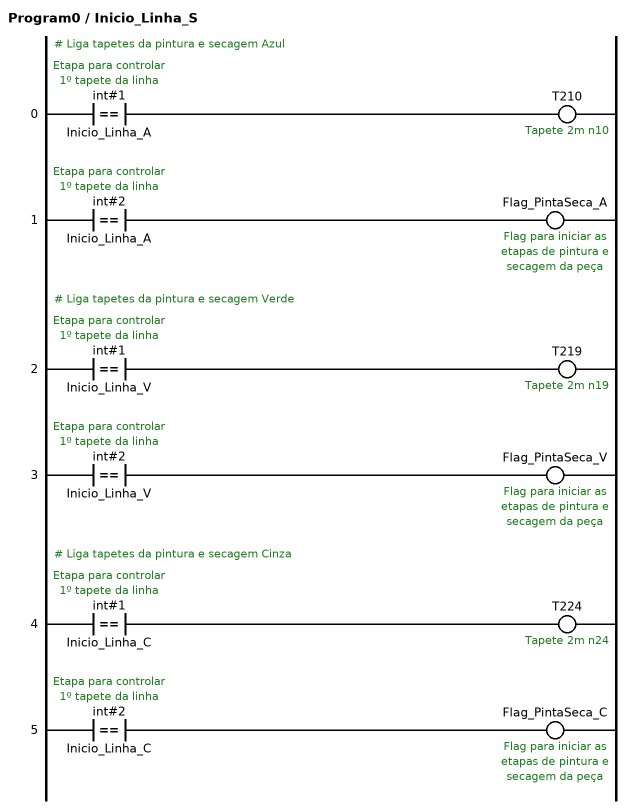
(* [picture p96: Program0 / Inicio_Linha_S, rungs 0-5] *)
(* Rung 0: # Liga tapetes da pintura e secagem Azul *)
T210 := int#1 = Inicio_Linha_A;
(* Rung 1 *)
Flag_PintaSeca_A := int#2 = Inicio_Linha_A;
(* Rung 2: # Liga tapetes da pintura e secagem Verde *)
T219 := int#1 = Inicio_Linha_V;
(* Rung 3 *)
Flag_PintaSeca_V := int#2 = Inicio_Linha_V;
(* Rung 4: # Liga tapetes da pintura e secagem Cinza *)
T224 := int#1 = Inicio_Linha_C;
(* Rung 5 *)
Flag_PintaSeca_C := int#2 = Inicio_Linha_C;

(* Section Pinta_Seca_E: ladder, written here as Structured Text *)

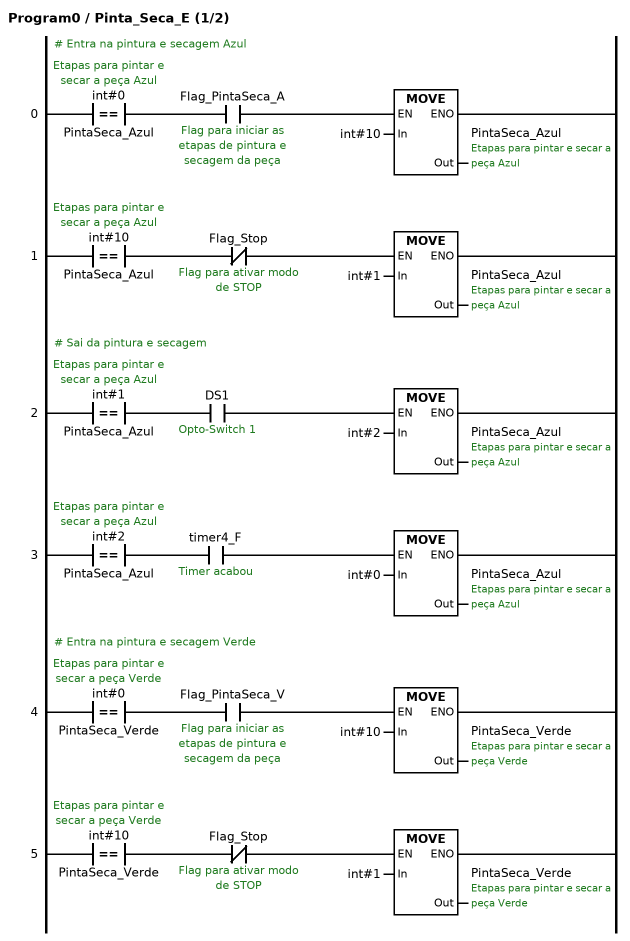
(* Rung 0: # Entra na pintura e secagem Azul *)
IF (int#0 = PintaSeca_Azul) AND Flag_PintaSeca_A THEN PintaSeca_Azul := int#10; END_IF;
(* Rung 1 *)
IF (int#10 = PintaSeca_Azul) AND NOT Flag_Stop THEN PintaSeca_Azul := int#1; END_IF;
(* Rung 2: # Sai da pintura e secagem *)
IF (int#1 = PintaSeca_Azul) AND DS1 THEN PintaSeca_Azul := int#2; END_IF;
(* Rung 3 *)
IF (int#2 = PintaSeca_Azul) AND timer4_F THEN PintaSeca_Azul := int#0; END_IF;
(* Rung 4: # Entra na pintura e secagem Verde *)
IF (int#0 = PintaSeca_Verde) AND Flag_PintaSeca_V THEN PintaSeca_Verde := int#10; END_IF;
(* Rung 5 *)
IF (int#10 = PintaSeca_Verde) AND NOT Flag_Stop THEN PintaSeca_Verde := int#1; END_IF;

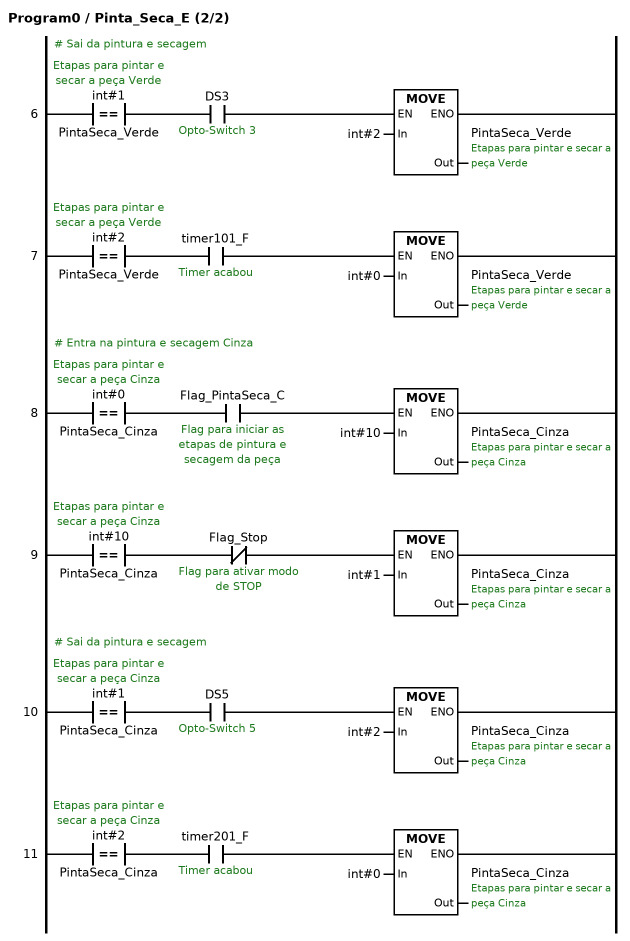
(* Rung 6: # Sai da pintura e secagem *)
IF (int#1 = PintaSeca_Verde) AND DS3 THEN PintaSeca_Verde := int#2; END_IF;
(* Rung 7 *)
IF (int#2 = PintaSeca_Verde) AND timer101_F THEN PintaSeca_Verde := int#0; END_IF;
(* Rung 8: # Entra na pintura e secagem Cinza *)
IF (int#0 = PintaSeca_Cinza) AND Flag_PintaSeca_C THEN PintaSeca_Cinza := int#10; END_IF;
(* Rung 9 *)
IF (int#10 = PintaSeca_Cinza) AND NOT Flag_Stop THEN PintaSeca_Cinza := int#1; END_IF;
(* Rung 10: # Sai da pintura e secagem *)
IF (int#1 = PintaSeca_Cinza) AND DS5 THEN PintaSeca_Cinza := int#2; END_IF;
(* Rung 11 *)
IF (int#2 = PintaSeca_Cinza) AND timer201_F THEN PintaSeca_Cinza := int#0; END_IF;

(* Section Pinta_Seca_S: ladder, written here as Structured Text *)

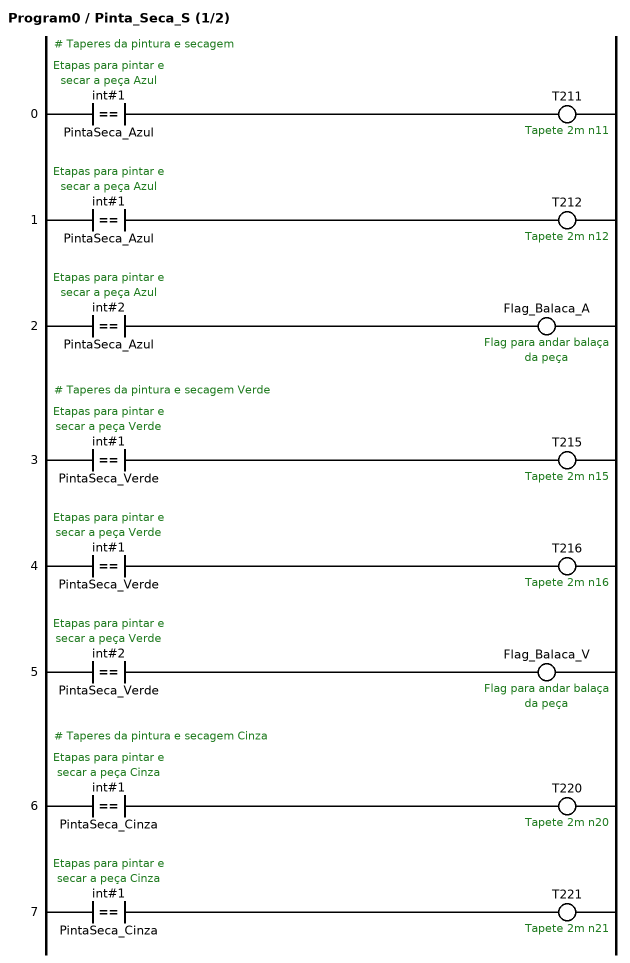
(* Rung 0: # Taperes da pintura e secagem *)
T211 := int#1 = PintaSeca_Azul;
(* Rung 1 *)
T212 := int#1 = PintaSeca_Azul;
(* Rung 2 *)
Flag_Balaca_A := int#2 = PintaSeca_Azul;
(* Rung 3: # Taperes da pintura e secagem Verde *)
T215 := int#1 = PintaSeca_Verde;
(* Rung 4 *)
T216 := int#1 = PintaSeca_Verde;
(* Rung 5 *)
Flag_Balaca_V := int#2 = PintaSeca_Verde;
(* Rung 6: # Taperes da pintura e secagem Cinza *)
T220 := int#1 = PintaSeca_Cinza;
(* Rung 7 *)
T221 := int#1 = PintaSeca_Cinza;

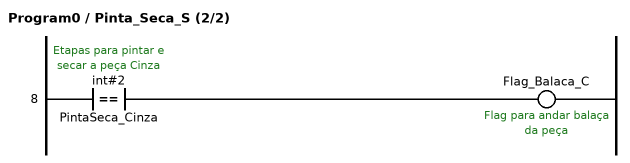
(* Rung 8 *)
Flag_Balaca_C := int#2 = PintaSeca_Cinza;

(* Section Balaca_E: ladder, written here as Structured Text *)

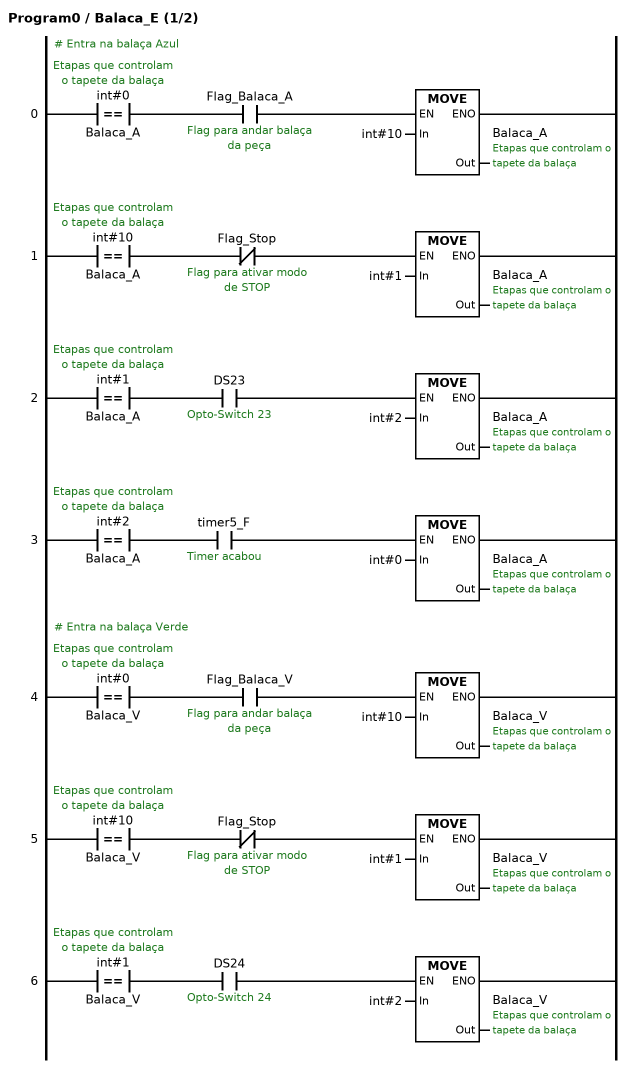
(* Rung 0: # Entra na balaça Azul *)
IF (int#0 = Balaca_A) AND Flag_Balaca_A THEN Balaca_A := int#10; END_IF;
(* Rung 1 *)
IF (int#10 = Balaca_A) AND NOT Flag_Stop THEN Balaca_A := int#1; END_IF;
(* Rung 2 *)
IF (int#1 = Balaca_A) AND DS23 THEN Balaca_A := int#2; END_IF;
(* Rung 3 *)
IF (int#2 = Balaca_A) AND timer5_F THEN Balaca_A := int#0; END_IF;
(* Rung 4: # Entra na balaça Verde *)
IF (int#0 = Balaca_V) AND Flag_Balaca_V THEN Balaca_V := int#10; END_IF;
(* Rung 5 *)
IF (int#10 = Balaca_V) AND NOT Flag_Stop THEN Balaca_V := int#1; END_IF;
(* Rung 6 *)
IF (int#1 = Balaca_V) AND DS24 THEN Balaca_V := int#2; END_IF;

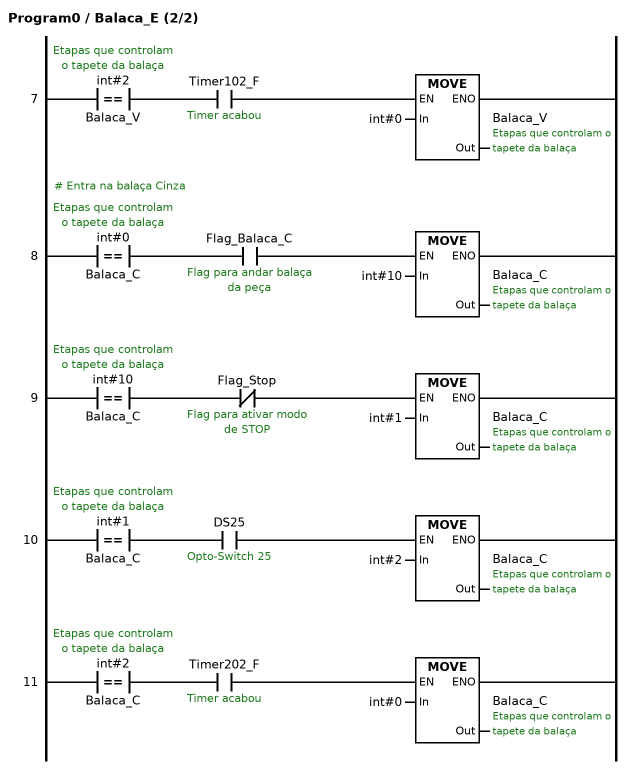
(* Rung 7 *)
IF (int#2 = Balaca_V) AND Timer102_F THEN Balaca_V := int#0; END_IF;
(* Rung 8: # Entra na balaça Cinza *)
IF (int#0 = Balaca_C) AND Flag_Balaca_C THEN Balaca_C := int#10; END_IF;
(* Rung 9 *)
IF (int#10 = Balaca_C) AND NOT Flag_Stop THEN Balaca_C := int#1; END_IF;
(* Rung 10 *)
IF (int#1 = Balaca_C) AND DS25 THEN Balaca_C := int#2; END_IF;
(* Rung 11 *)
IF (int#2 = Balaca_C) AND Timer202_F THEN Balaca_C := int#0; END_IF;

(* Section Balaca_S: ladder, written here as Structured Text *)

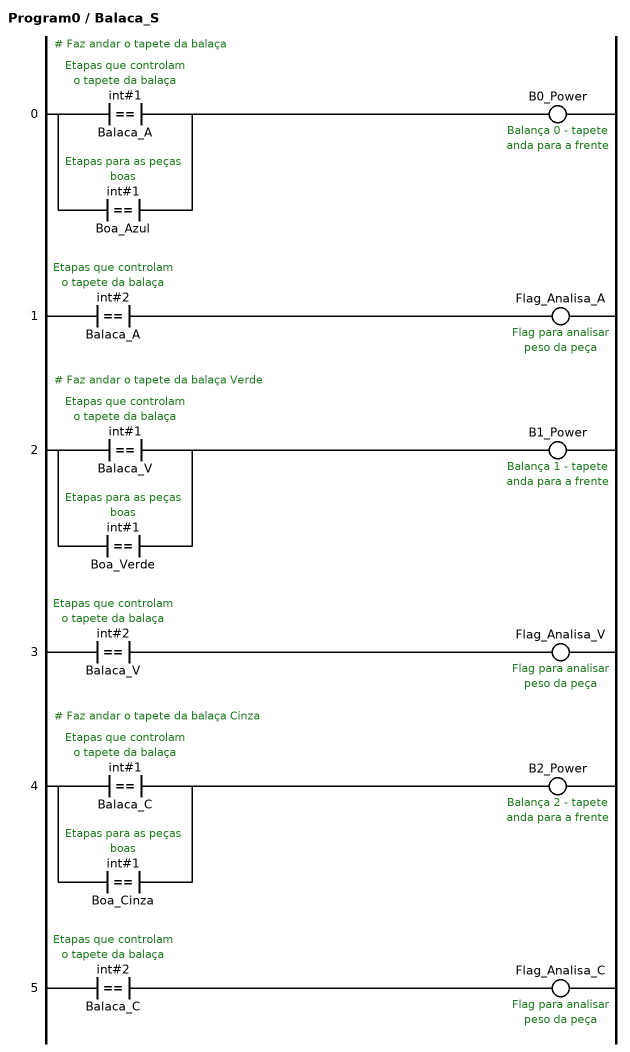
(* Rung 0: # Faz andar o tapete da balaça *)
B0_Power := (int#1 = Balaca_A) OR (int#1 = Boa_Azul);
(* Rung 1 *)
Flag_Analisa_A := int#2 = Balaca_A;
(* Rung 2: # Faz andar o tapete da balaça Verde *)
B1_Power := (int#1 = Balaca_V) OR (int#1 = Boa_Verde);
(* Rung 3 *)
Flag_Analisa_V := int#2 = Balaca_V;
(* Rung 4: # Faz andar o tapete da balaça Cinza *)
B2_Power := (int#1 = Balaca_C) OR (int#1 = Boa_Cinza);
(* Rung 5 *)
Flag_Analisa_C := int#2 = Balaca_C;

(* Section Analisa_Pesos_E: ladder, written here as Structured Text *)

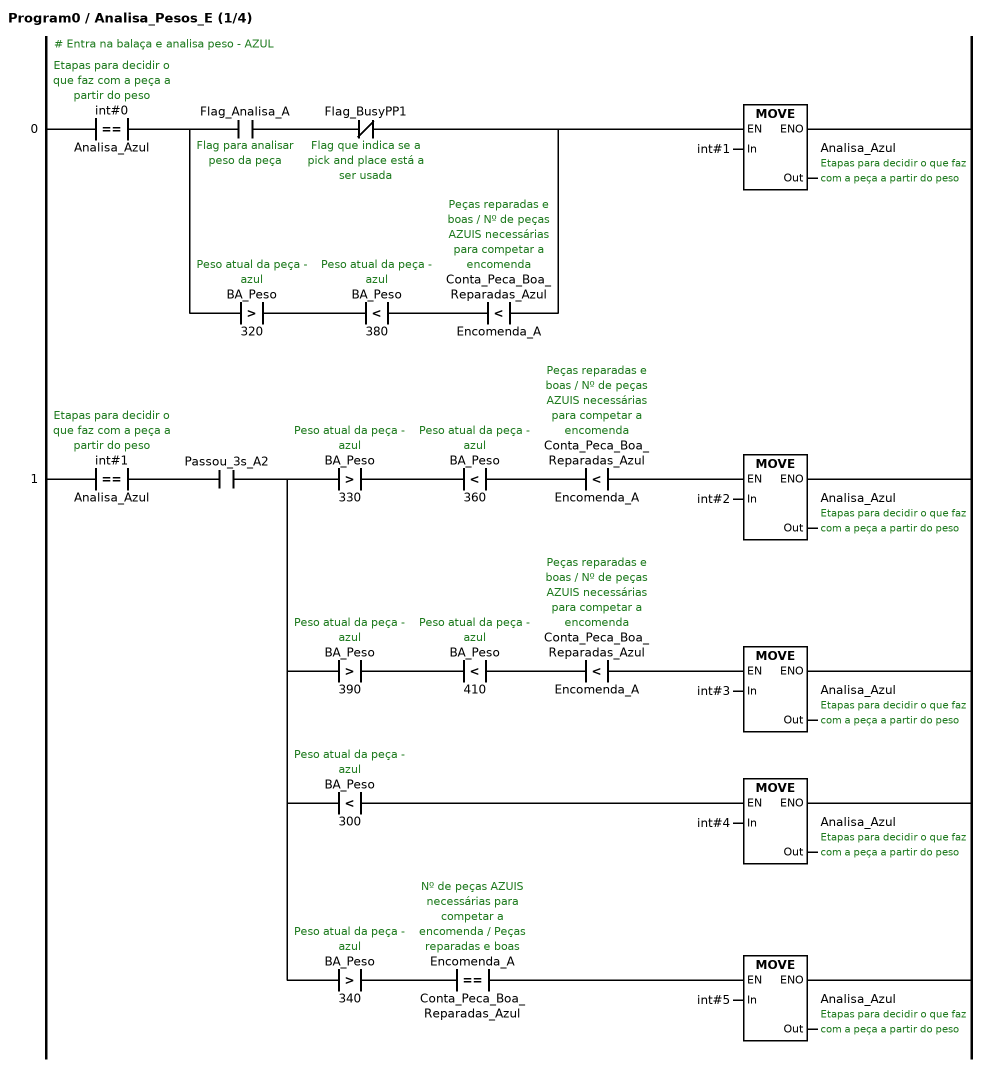
(* Rung 0: # Entra na balaça e analisa peso - AZUL *)
IF (int#0 = Analisa_Azul) AND ((Flag_Analisa_A AND NOT Flag_BusyPP1) OR ((BA_Peso > 320) AND (BA_Peso < 380) AND (Conta_Peca_Boa_Reparadas_Azul < Encomenda_A))) THEN
    Analisa_Azul := int#1;
END_IF;
(* Rung 1 *)
_p32 := (int#1 = Analisa_Azul) AND Passou_3s_A2;
IF (int#1 = Analisa_Azul) AND Passou_3s_A2 AND (BA_Peso > 330) AND (BA_Peso < 360) AND (Conta_Peca_Boa_Reparadas_Azul < Encomenda_A) THEN
    Analisa_Azul := int#2;
END_IF;
IF _p32 AND (BA_Peso > 390) AND (BA_Peso < 410) AND (Conta_Peca_Boa_Reparadas_Azul < Encomenda_A) THEN
    Analisa_Azul := int#3;
END_IF;
IF _p32 AND (BA_Peso < 300) THEN Analisa_Azul := int#4; END_IF;
IF _p32 AND (BA_Peso > 340) AND (Encomenda_A = Conta_Peca_Boa_Reparadas_Azul) THEN
    Analisa_Azul := int#5;
END_IF;

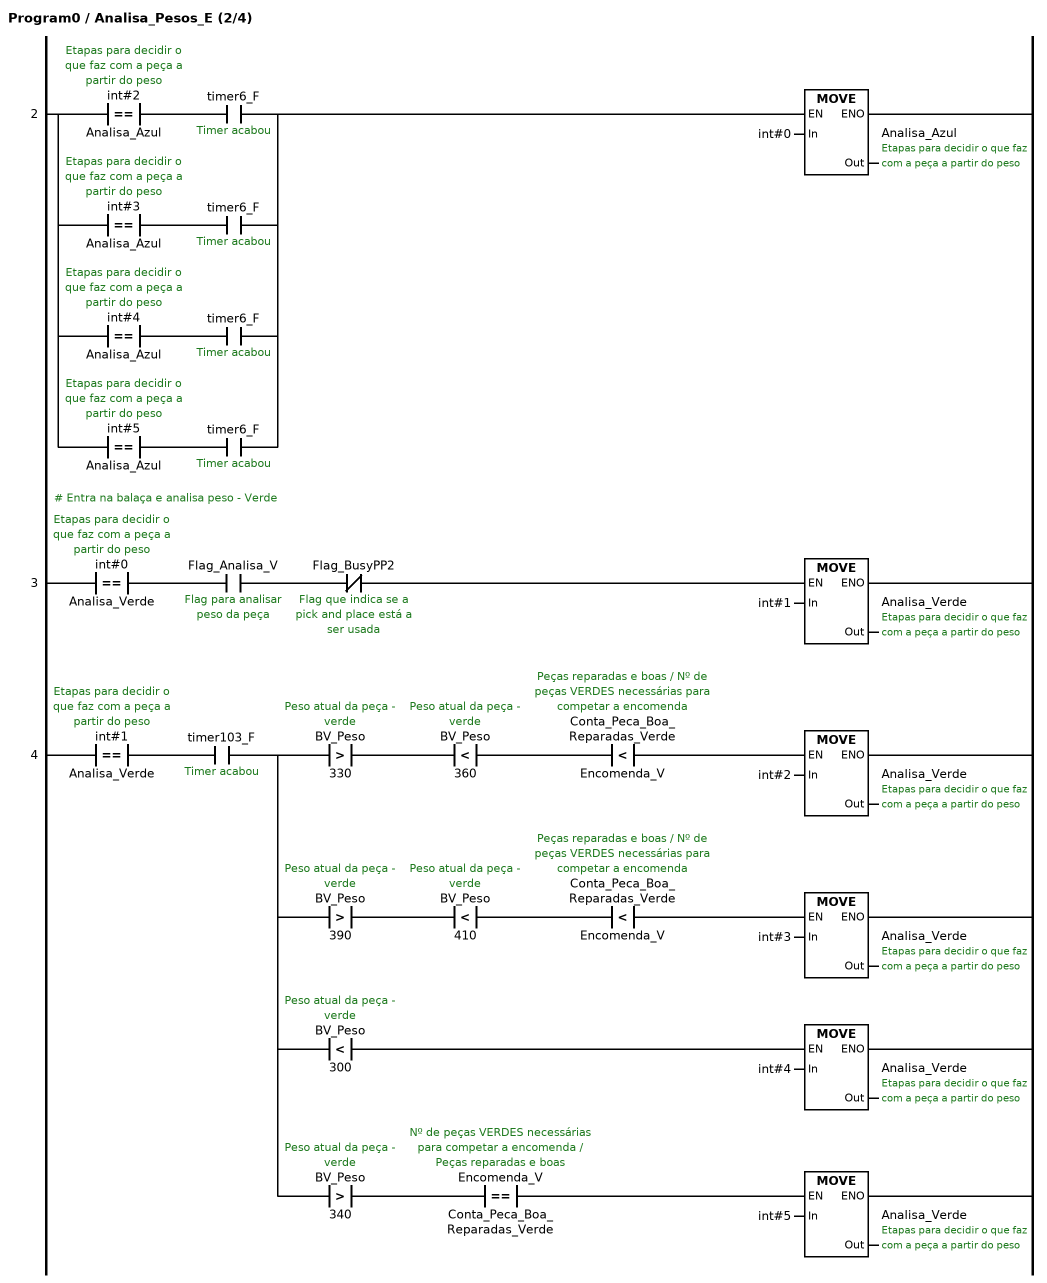
(* Rung 2 *)
IF ((int#2 = Analisa_Azul) AND timer6_F) OR ((int#3 = Analisa_Azul) AND timer6_F) OR ((int#4 = Analisa_Azul) AND timer6_F) OR ((int#5 = Analisa_Azul) AND timer6_F) THEN
    Analisa_Azul := int#0;
END_IF;
(* Rung 3: # Entra na balaça e analisa peso - Verde *)
IF (int#0 = Analisa_Verde) AND Flag_Analisa_V AND NOT Flag_BusyPP2 THEN Analisa_Verde := int#1; END_IF;
(* Rung 4 *)
_p33 := (int#1 = Analisa_Verde) AND timer103_F;
IF (int#1 = Analisa_Verde) AND timer103_F AND (BV_Peso > 330) AND (BV_Peso < 360) AND (Conta_Peca_Boa_Reparadas_Verde < Encomenda_V) THEN
    Analisa_Verde := int#2;
END_IF;
IF _p33 AND (BV_Peso > 390) AND (BV_Peso < 410) AND (Conta_Peca_Boa_Reparadas_Verde < Encomenda_V) THEN
    Analisa_Verde := int#3;
END_IF;
IF _p33 AND (BV_Peso < 300) THEN Analisa_Verde := int#4; END_IF;
IF _p33 AND (BV_Peso > 340) AND (Encomenda_V = Conta_Peca_Boa_Reparadas_Verde) THEN
    Analisa_Verde := int#5;
END_IF;

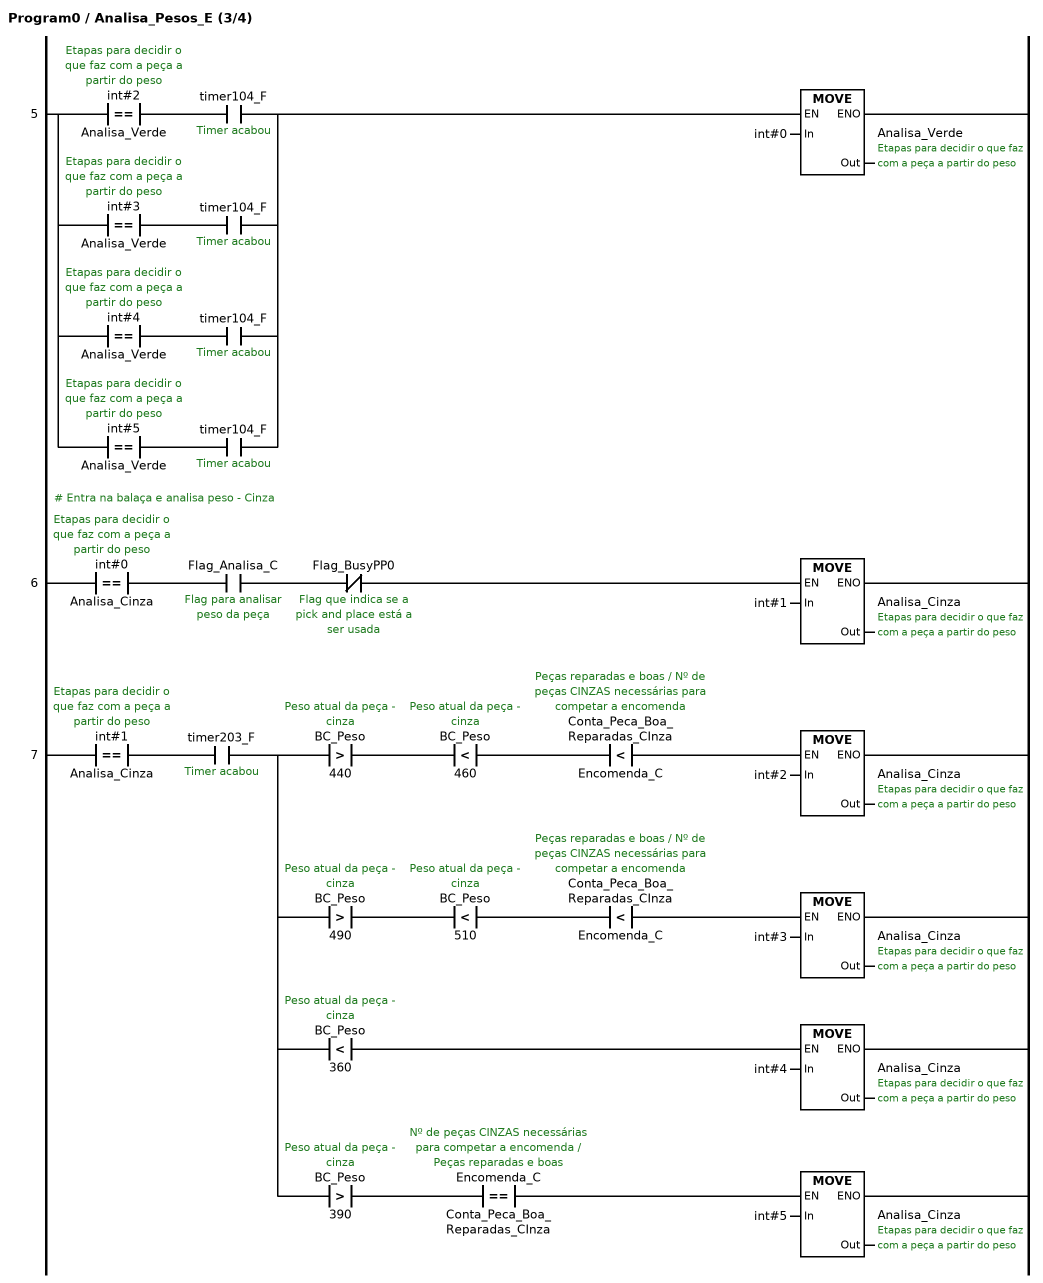
(* Rung 5 *)
IF ((int#2 = Analisa_Verde) AND timer104_F) OR ((int#3 = Analisa_Verde) AND timer104_F) OR ((int#4 = Analisa_Verde) AND timer104_F) OR ((int#5 = Analisa_Verde) AND timer104_F) THEN
    Analisa_Verde := int#0;
END_IF;
(* Rung 6: # Entra na balaça e analisa peso - Cinza *)
IF (int#0 = Analisa_Cinza) AND Flag_Analisa_C AND NOT Flag_BusyPP0 THEN Analisa_Cinza := int#1; END_IF;
(* Rung 7 *)
_p34 := (int#1 = Analisa_Cinza) AND timer203_F;
IF (int#1 = Analisa_Cinza) AND timer203_F AND (BC_Peso > 440) AND (BC_Peso < 460) AND (Conta_Peca_Boa_Reparadas_CInza < Encomenda_C) THEN
    Analisa_Cinza := int#2;
END_IF;
IF _p34 AND (BC_Peso > 490) AND (BC_Peso < 510) AND (Conta_Peca_Boa_Reparadas_CInza < Encomenda_C) THEN
    Analisa_Cinza := int#3;
END_IF;
IF _p34 AND (BC_Peso < 360) THEN Analisa_Cinza := int#4; END_IF;
IF _p34 AND (BC_Peso > 390) AND (Encomenda_C = Conta_Peca_Boa_Reparadas_CInza) THEN
    Analisa_Cinza := int#5;
END_IF;

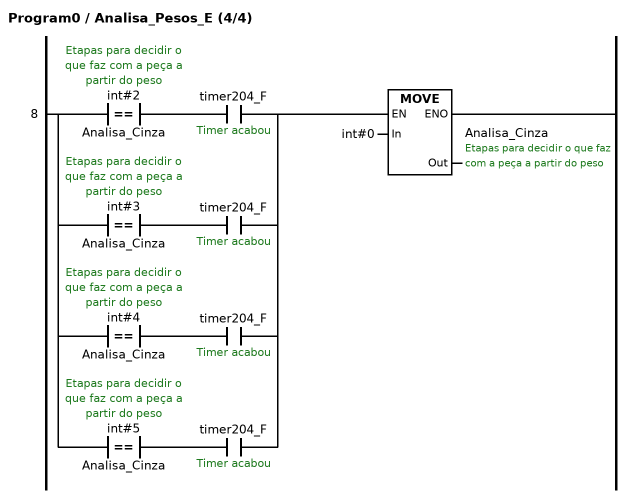
(* Rung 8 *)
IF ((int#2 = Analisa_Cinza) AND timer204_F) OR ((int#3 = Analisa_Cinza) AND timer204_F) OR ((int#4 = Analisa_Cinza) AND timer204_F) OR ((int#5 = Analisa_Cinza) AND timer204_F) THEN
    Analisa_Cinza := int#0;
END_IF;

(* Section Analisa_Pesos_S: ladder, written here as Structured Text *)

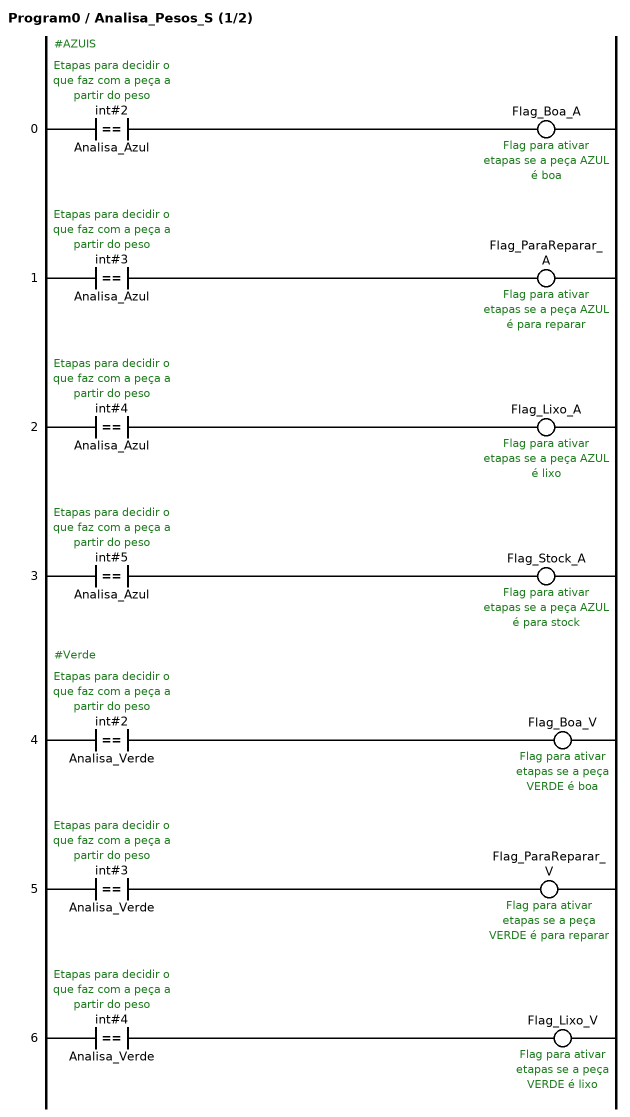
(* Rung 0: #AZUIS *)
Flag_Boa_A := int#2 = Analisa_Azul;
(* Rung 1 *)
Flag_ParaReparar_A := int#3 = Analisa_Azul;
(* Rung 2 *)
Flag_Lixo_A := int#4 = Analisa_Azul;
(* Rung 3 *)
Flag_Stock_A := int#5 = Analisa_Azul;
(* Rung 4: #Verde *)
Flag_Boa_V := int#2 = Analisa_Verde;
(* Rung 5 *)
Flag_ParaReparar_V := int#3 = Analisa_Verde;
(* Rung 6 *)
Flag_Lixo_V := int#4 = Analisa_Verde;

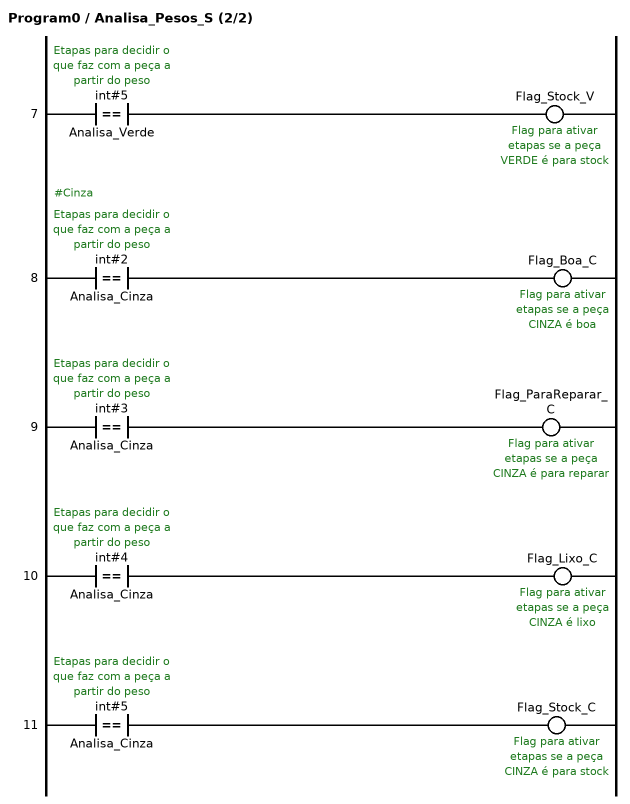
(* Rung 7 *)
Flag_Stock_V := int#5 = Analisa_Verde;
(* Rung 8: #Cinza *)
Flag_Boa_C := int#2 = Analisa_Cinza;
(* Rung 9 *)
Flag_ParaReparar_C := int#3 = Analisa_Cinza;
(* Rung 10 *)
Flag_Lixo_C := int#4 = Analisa_Cinza;
(* Rung 11 *)
Flag_Stock_C := int#5 = Analisa_Cinza;

(* Section Boas_E: ladder, written here as Structured Text *)

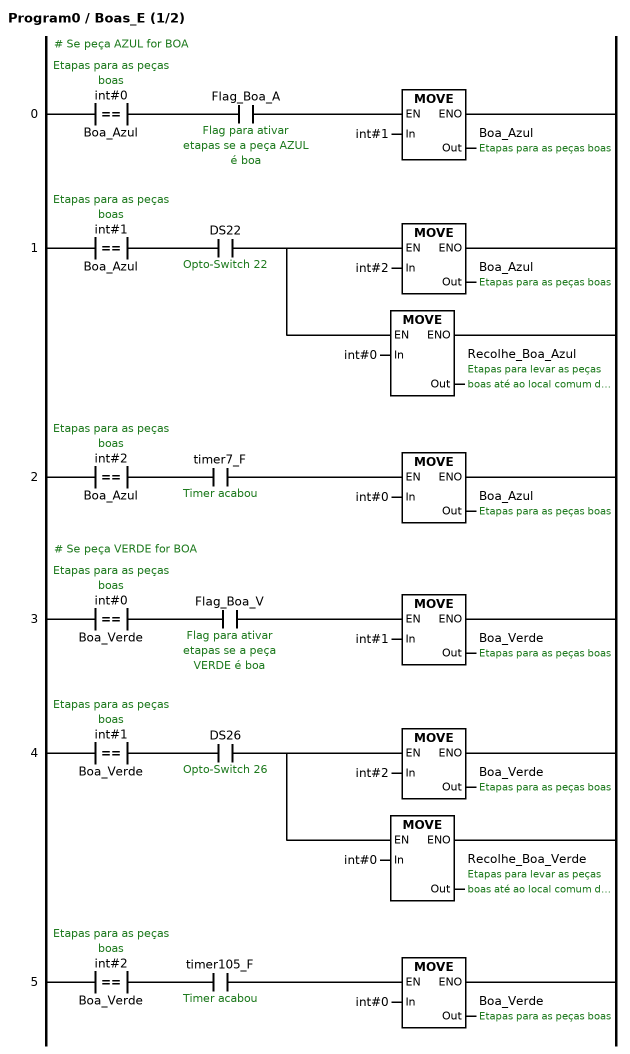
(* Rung 0: # Se peça AZUL for BOA *)
IF (int#0 = Boa_Azul) AND Flag_Boa_A THEN Boa_Azul := int#1; END_IF;
(* Rung 1 *)
_p35 := (int#1 = Boa_Azul) AND DS22;
IF _p35 THEN
    Boa_Azul := int#2;
    Recolhe_Boa_Azul := int#0;
END_IF;
(* Rung 2 *)
IF (int#2 = Boa_Azul) AND timer7_F THEN Boa_Azul := int#0; END_IF;
(* Rung 3: # Se peça VERDE for BOA *)
IF (int#0 = Boa_Verde) AND Flag_Boa_V THEN Boa_Verde := int#1; END_IF;
(* Rung 4 *)
_p36 := (int#1 = Boa_Verde) AND DS26;
IF _p36 THEN
    Boa_Verde := int#2;
    Recolhe_Boa_Verde := int#0;
END_IF;
(* Rung 5 *)
IF (int#2 = Boa_Verde) AND timer105_F THEN Boa_Verde := int#0; END_IF;

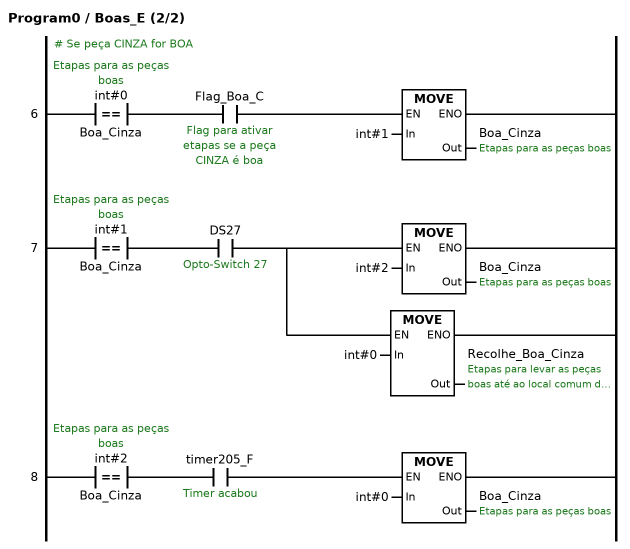
(* Rung 6: # Se peça CINZA for BOA *)
IF (int#0 = Boa_Cinza) AND Flag_Boa_C THEN Boa_Cinza := int#1; END_IF;
(* Rung 7 *)
_p37 := (int#1 = Boa_Cinza) AND DS27;
IF _p37 THEN
    Boa_Cinza := int#2;
    Recolhe_Boa_Cinza := int#0;
END_IF;
(* Rung 8 *)
IF (int#2 = Boa_Cinza) AND timer205_F THEN Boa_Cinza := int#0; END_IF;

(* Section Boas_S: ladder, written here as Structured Text *)

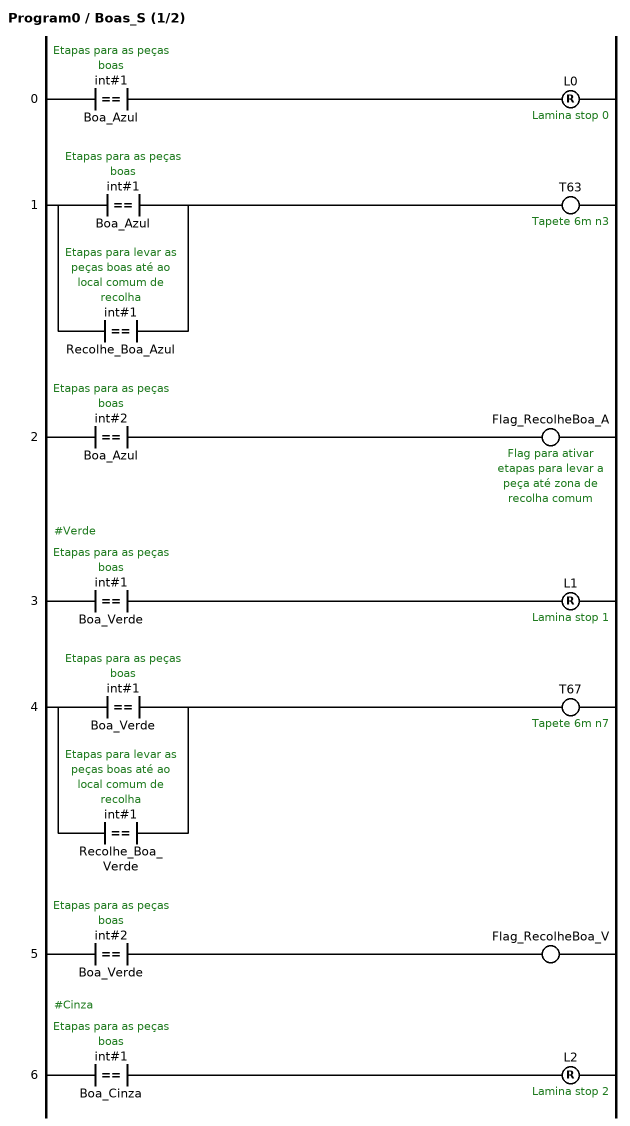
(* Rung 0 *)
IF int#1 = Boa_Azul THEN L0 := FALSE; END_IF;
(* Rung 1 *)
T63 := (int#1 = Boa_Azul) OR (int#1 = Recolhe_Boa_Azul);
(* Rung 2 *)
Flag_RecolheBoa_A := int#2 = Boa_Azul;
(* Rung 3: #Verde *)
IF int#1 = Boa_Verde THEN L1 := FALSE; END_IF;
(* Rung 4 *)
T67 := (int#1 = Boa_Verde) OR (int#1 = Recolhe_Boa_Verde);
(* Rung 5 *)
Flag_RecolheBoa_V := int#2 = Boa_Verde;
(* Rung 6: #Cinza *)
IF int#1 = Boa_Cinza THEN L2 := FALSE; END_IF;

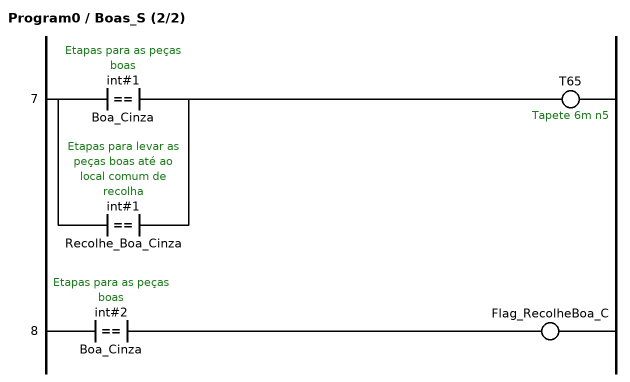
(* Rung 7 *)
T65 := (int#1 = Boa_Cinza) OR (int#1 = Recolhe_Boa_Cinza);
(* Rung 8 *)
Flag_RecolheBoa_C := int#2 = Boa_Cinza;

(* Section Recolhe_Boa_E: ladder, written here as Structured Text *)

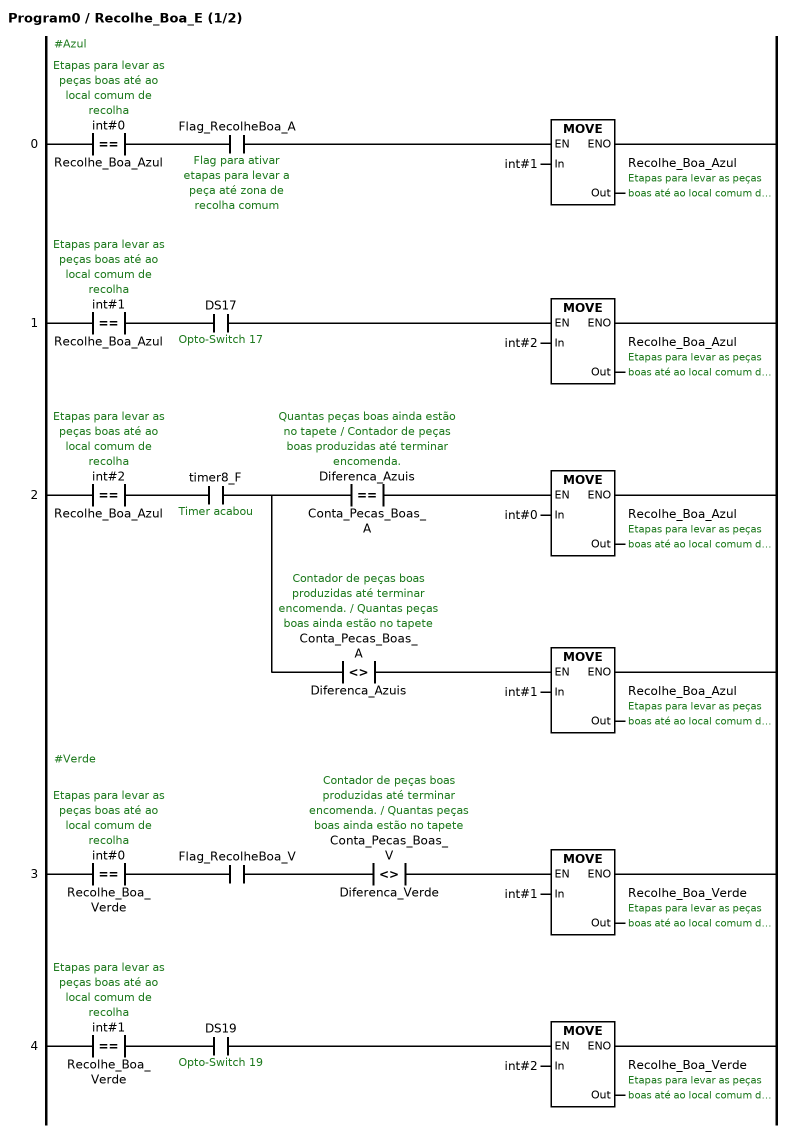
(* Rung 0: #Azul *)
IF (int#0 = Recolhe_Boa_Azul) AND Flag_RecolheBoa_A THEN Recolhe_Boa_Azul := int#1; END_IF;
(* Rung 1 *)
IF (int#1 = Recolhe_Boa_Azul) AND DS17 THEN Recolhe_Boa_Azul := int#2; END_IF;
(* Rung 2 *)
_p38 := (int#2 = Recolhe_Boa_Azul) AND timer8_F;
IF (int#2 = Recolhe_Boa_Azul) AND timer8_F AND (Diferenca_Azuis = Conta_Pecas_Boas_A) THEN
    Recolhe_Boa_Azul := int#0;
END_IF;
IF _p38 AND (Conta_Pecas_Boas_A <> Diferenca_Azuis) THEN Recolhe_Boa_Azul := int#1; END_IF;
(* Rung 3: #Verde *)
IF (int#0 = Recolhe_Boa_Verde) AND Flag_RecolheBoa_V AND (Conta_Pecas_Boas_V <> Diferenca_Verde) THEN
    Recolhe_Boa_Verde := int#1;
END_IF;
(* Rung 4 *)
IF (int#1 = Recolhe_Boa_Verde) AND DS19 THEN Recolhe_Boa_Verde := int#2; END_IF;

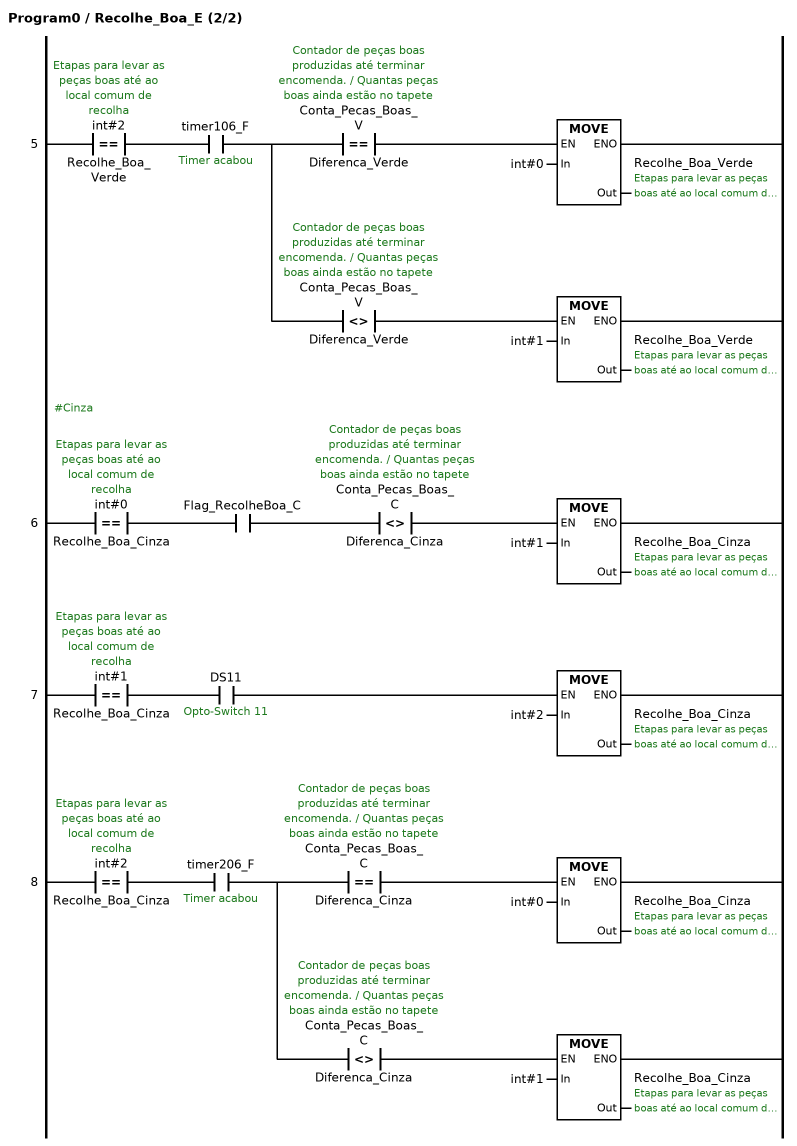
(* Rung 5 *)
_p39 := (int#2 = Recolhe_Boa_Verde) AND timer106_F;
IF (int#2 = Recolhe_Boa_Verde) AND timer106_F AND (Conta_Pecas_Boas_V = Diferenca_Verde) THEN
    Recolhe_Boa_Verde := int#0;
END_IF;
IF _p39 AND (Conta_Pecas_Boas_V <> Diferenca_Verde) THEN Recolhe_Boa_Verde := int#1; END_IF;
(* Rung 6: #Cinza *)
IF (int#0 = Recolhe_Boa_Cinza) AND Flag_RecolheBoa_C AND (Conta_Pecas_Boas_C <> Diferenca_Cinza) THEN
    Recolhe_Boa_Cinza := int#1;
END_IF;
(* Rung 7 *)
IF (int#1 = Recolhe_Boa_Cinza) AND DS11 THEN Recolhe_Boa_Cinza := int#2; END_IF;
(* Rung 8 *)
_p40 := (int#2 = Recolhe_Boa_Cinza) AND timer206_F;
IF (int#2 = Recolhe_Boa_Cinza) AND timer206_F AND (Conta_Pecas_Boas_C = Diferenca_Cinza) THEN
    Recolhe_Boa_Cinza := int#0;
END_IF;
IF _p40 AND (Conta_Pecas_Boas_C <> Diferenca_Cinza) THEN Recolhe_Boa_Cinza := int#1; END_IF;

(* Section Recolhe_Boa_S: ladder, written here as Structured Text *)

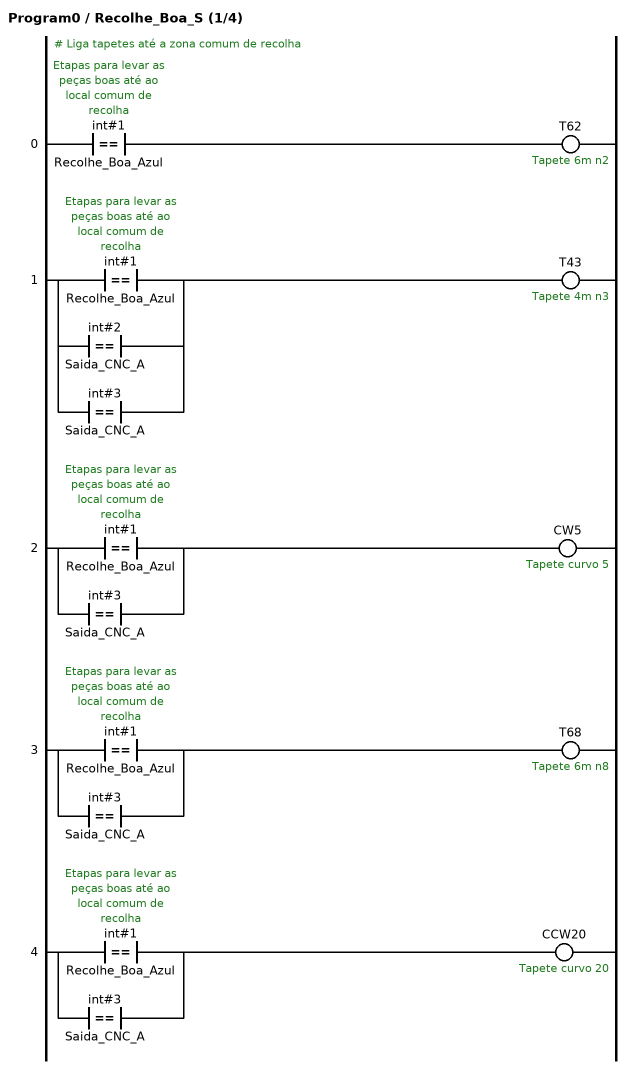
(* Rung 0: # Liga tapetes até a zona comum de recolha *)
T62 := int#1 = Recolhe_Boa_Azul;
(* Rung 1 *)
T43 := (int#1 = Recolhe_Boa_Azul) OR (int#2 = Saida_CNC_A) OR (int#3 = Saida_CNC_A);
(* Rung 2 *)
CW5 := (int#1 = Recolhe_Boa_Azul) OR (int#3 = Saida_CNC_A);
(* Rung 3 *)
T68 := (int#1 = Recolhe_Boa_Azul) OR (int#3 = Saida_CNC_A);
(* Rung 4 *)
CCW20 := (int#1 = Recolhe_Boa_Azul) OR (int#3 = Saida_CNC_A);

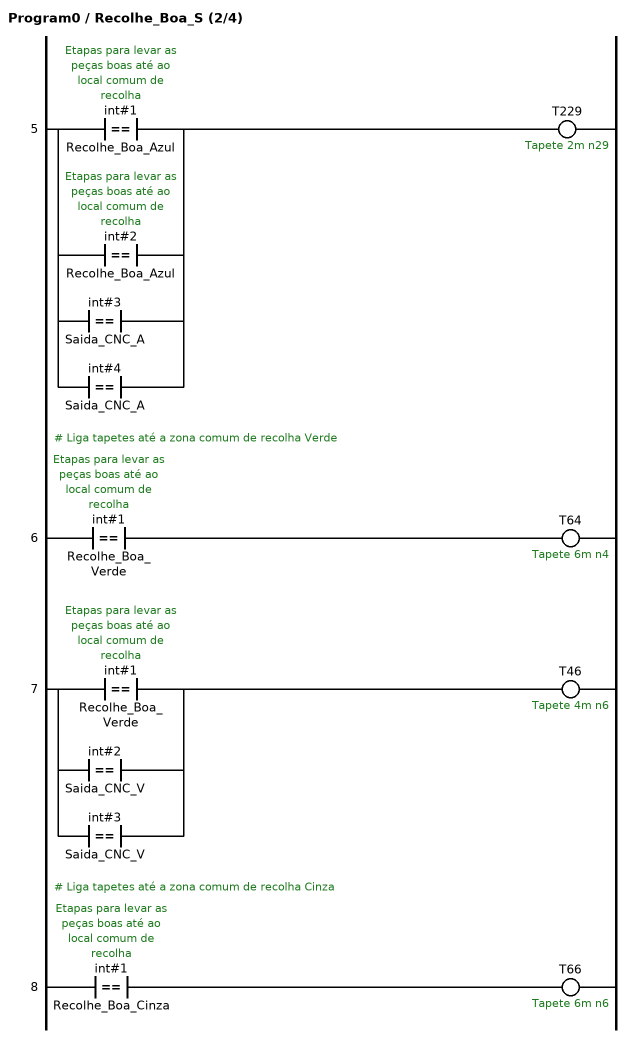
(* Rung 5 *)
T229 := (int#1 = Recolhe_Boa_Azul) OR (int#2 = Recolhe_Boa_Azul) OR (int#3 = Saida_CNC_A) OR (int#4 = Saida_CNC_A);
(* Rung 6: # Liga tapetes até a zona comum de recolha Verde *)
T64 := int#1 = Recolhe_Boa_Verde;
(* Rung 7 *)
T46 := (int#1 = Recolhe_Boa_Verde) OR (int#2 = Saida_CNC_V) OR (int#3 = Saida_CNC_V);
(* Rung 8: # Liga tapetes até a zona comum de recolha Cinza *)
T66 := int#1 = Recolhe_Boa_Cinza;

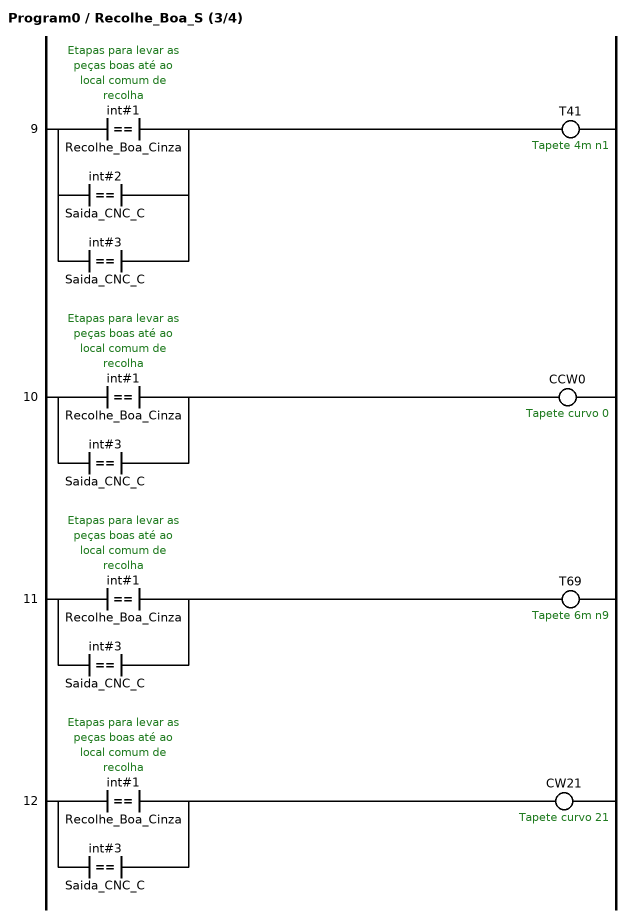
(* Rung 9 *)
T41 := (int#1 = Recolhe_Boa_Cinza) OR (int#2 = Saida_CNC_C) OR (int#3 = Saida_CNC_C);
(* Rung 10 *)
CCW0 := (int#1 = Recolhe_Boa_Cinza) OR (int#3 = Saida_CNC_C);
(* Rung 11 *)
T69 := (int#1 = Recolhe_Boa_Cinza) OR (int#3 = Saida_CNC_C);
(* Rung 12 *)
CW21 := (int#1 = Recolhe_Boa_Cinza) OR (int#3 = Saida_CNC_C);

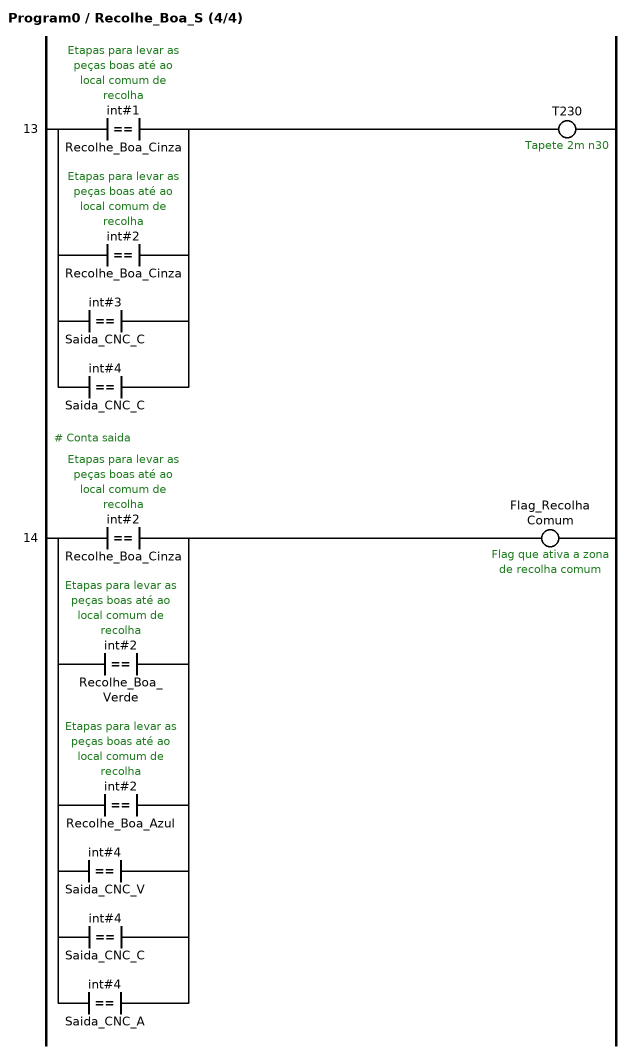
(* Rung 13 *)
T230 := (int#1 = Recolhe_Boa_Cinza) OR (int#2 = Recolhe_Boa_Cinza) OR (int#3 = Saida_CNC_C) OR (int#4 = Saida_CNC_C);
(* Rung 14: # Conta saida *)
Flag_RecolhaComum := (int#2 = Recolhe_Boa_Cinza) OR (int#2 = Recolhe_Boa_Verde) OR (int#2 = Recolhe_Boa_Azul) OR (int#4 = Saida_CNC_V) OR (int#4 = Saida_CNC_C) OR (int#4 = Saida_CNC_A);

(* Section Lixo_E: ladder, written here as Structured Text *)

